(* Schneider Machine Expert - Basic project m200-cpp EXPERIMENTAL, file version 3.0.0.0 *)
(* ProjectInformations: Name=New project *)

HARDWARE
  Cpu 0: TM200CE40T
  EthernetConfiguration: NetworkName=M200, IpAllocationMode=FixedAddress, IpAddress=0.0.0.0, SubnetMask=0.0.0.0
  SerialLineConfiguration: Baud=Baud19200, Parity=ParityEven, DataBits=DataBits8, StopBits=StopBits1, PhysicalMedium=PhysicalMediumRs485, TransmissionMode=TransmissionModeModbusRtu, SlaveId=1, Addressing=SlaveAddressing
  MastTask: UsePeriodScanMode=false, PeriodScan=100
  FastTask: Period=255
  CpuBehavior: StartingMode=StartAsPreviousState, AutoSaveRamOnEeprom=true, WatchdogPeriod=250

SYMBOLS  (address, symbol, comment, settings)
  %S13      SB_FIRSTRUN  "Indicates the first controller cycle in RUN mode"
  %R0         [Type=Fifo]
  %M0       compiler_reused_M0_0
  %M1       compiler_reused_M1_1
  %M2       compiler_reused_M2_2
  %M3       compiler_reused_M3_3

POU Generated C++ - EXPERIMENTAL
  (* SectionNumber=0 *)

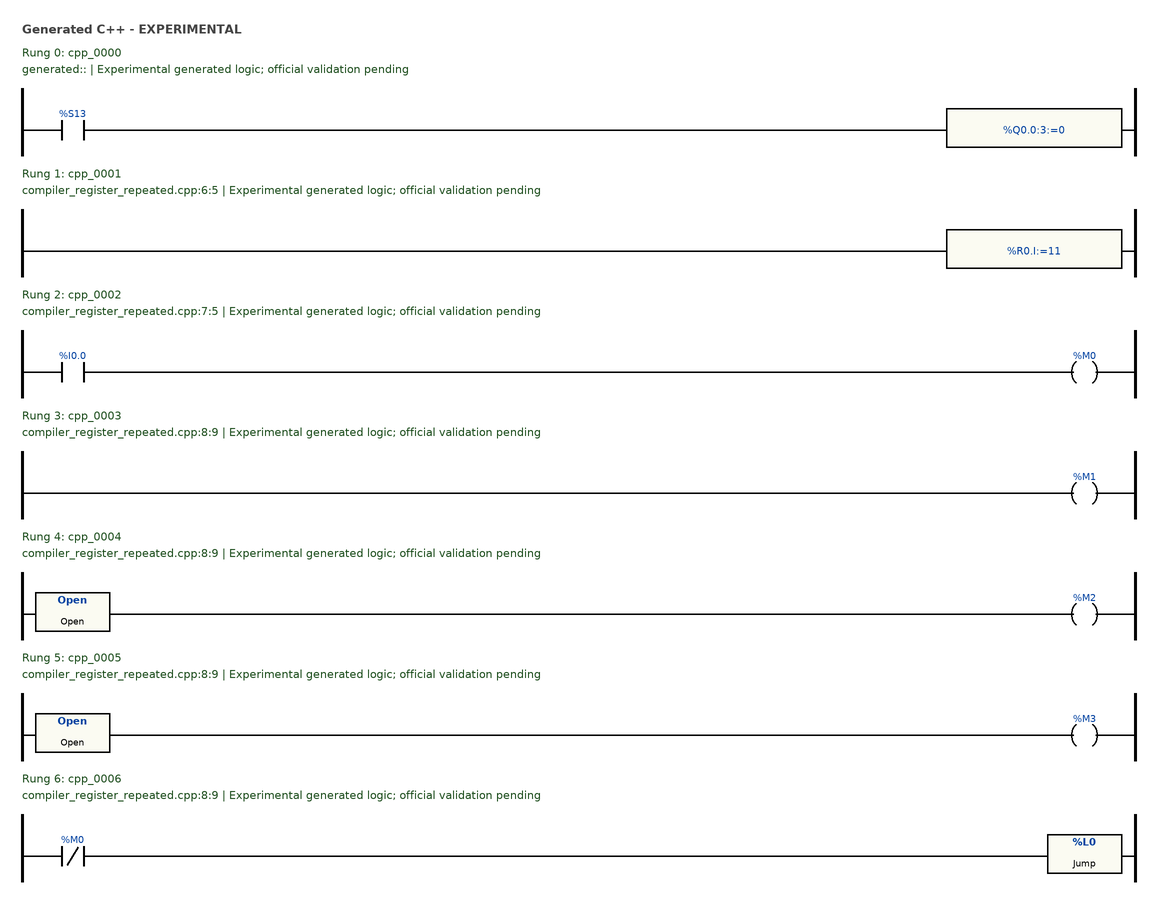

// Rung 0: cpp_0000
// generated:: | Experimental generated logic; official validation pending
  LD %S13                 (* SB_FIRSTRUN *)
  [%Q0.0:3:=0]
  // as ST:
  //   IF SB_FIRSTRUN THEN %Q0.0:3:=0; END_IF;

// Rung 1: cpp_0001
// compiler_register_repeated.cpp:6:5 | Experimental generated logic; official validation pending
  LD 1
  [%R0.I:=11]
  // as ST:
  //   %R0.I:=11;

// Rung 2: cpp_0002
// compiler_register_repeated.cpp:7:5 | Experimental generated logic; official validation pending
  LD %I0.0
  ST %M0                  (* compiler_reused_M0_0 *)
  // as ST:
  //   compiler_reused_M0_0 := %I0.0;

// Rung 3: cpp_0003
// compiler_register_repeated.cpp:8:9 | Experimental generated logic; official validation pending
  LD 1
  ST %M1                  (* compiler_reused_M1_1 *)
  // as ST:
  //   compiler_reused_M1_1 := TRUE;

// Rung 4: cpp_0004
// compiler_register_repeated.cpp:8:9 | Experimental generated logic; official validation pending
  LD 0
  ST %M2                  (* compiler_reused_M2_2 *)
  // as ST:
  //   compiler_reused_M2_2 := FALSE;

// Rung 5: cpp_0005
// compiler_register_repeated.cpp:8:9 | Experimental generated logic; official validation pending
  LD 0
  ST %M3                  (* compiler_reused_M3_3 *)
  // as ST:
  //   compiler_reused_M3_3 := FALSE;

// Rung 6: cpp_0006
// compiler_register_repeated.cpp:8:9 | Experimental generated logic; official validation pending
  LDN %M0                 (* compiler_reused_M0_0 *)
  JMPC %L0
  // as ST:
  //   IF NOT compiler_reused_M0_0 THEN JMP %L0; END_IF;

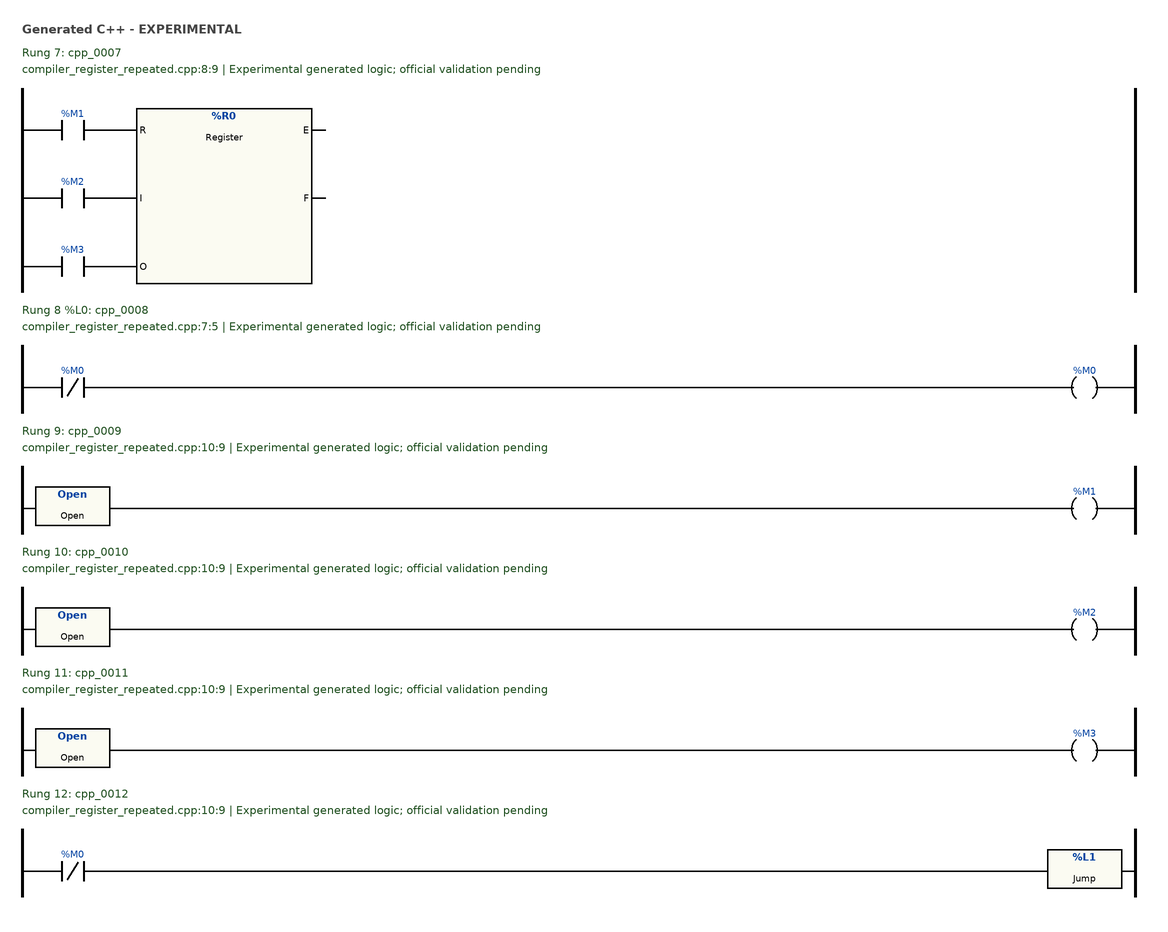

// Rung 7: cpp_0007
// compiler_register_repeated.cpp:8:9 | Experimental generated logic; official validation pending
  BLK %R0
  LD %M1                  (* compiler_reused_M1_1 *)
  R
  LD %M2                  (* compiler_reused_M2_2 *)
  I
  LD %M3                  (* compiler_reused_M3_3 *)
  O
  END_BLK
  // as ST:
  //   %R0(R := compiler_reused_M1_1, I := compiler_reused_M2_2, O := compiler_reused_M3_3);

// Rung 8 %L0: cpp_0008
// compiler_register_repeated.cpp:7:5 | Experimental generated logic; official validation pending
  %L0:
  LDN %M0                 (* compiler_reused_M0_0 *)
  ST %M0                  (* compiler_reused_M0_0 *)
  // as ST:
  //   %L0:
  //   compiler_reused_M0_0 := NOT compiler_reused_M0_0;

// Rung 9: cpp_0009
// compiler_register_repeated.cpp:10:9 | Experimental generated logic; official validation pending
  LD 0
  ST %M1                  (* compiler_reused_M1_1 *)
  // as ST:
  //   compiler_reused_M1_1 := FALSE;

// Rung 10: cpp_0010
// compiler_register_repeated.cpp:10:9 | Experimental generated logic; official validation pending
  LD 0
  ST %M2                  (* compiler_reused_M2_2 *)
  // as ST:
  //   compiler_reused_M2_2 := FALSE;

// Rung 11: cpp_0011
// compiler_register_repeated.cpp:10:9 | Experimental generated logic; official validation pending
  LD 0
  ST %M3                  (* compiler_reused_M3_3 *)
  // as ST:
  //   compiler_reused_M3_3 := FALSE;

// Rung 12: cpp_0012
// compiler_register_repeated.cpp:10:9 | Experimental generated logic; official validation pending
  LDN %M0                 (* compiler_reused_M0_0 *)
  JMPC %L1
  // as ST:
  //   IF NOT compiler_reused_M0_0 THEN JMP %L1; END_IF;

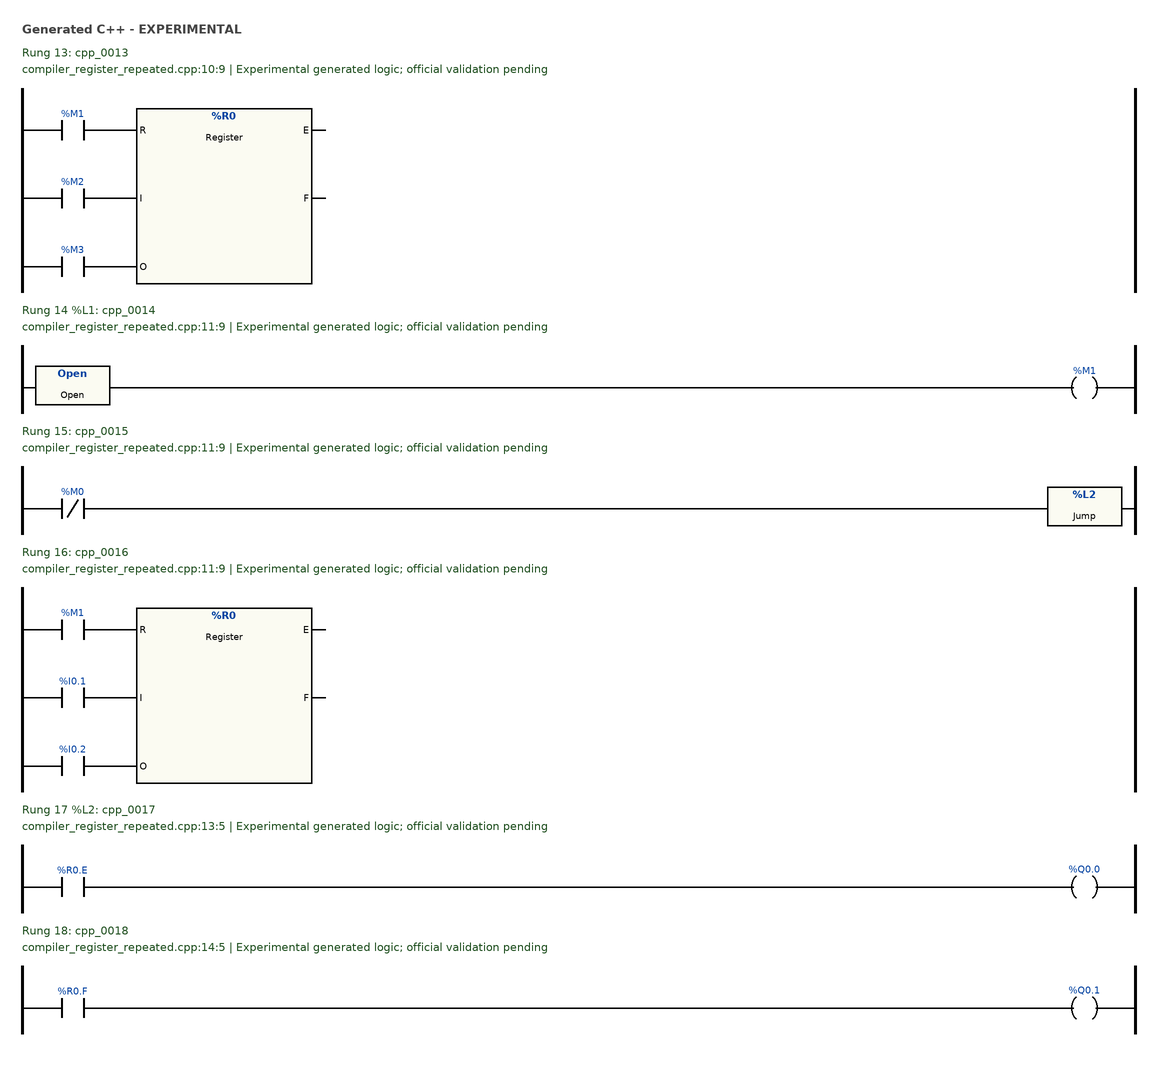

// Rung 13: cpp_0013
// compiler_register_repeated.cpp:10:9 | Experimental generated logic; official validation pending
  BLK %R0
  LD %M1                  (* compiler_reused_M1_1 *)
  R
  LD %M2                  (* compiler_reused_M2_2 *)
  I
  LD %M3                  (* compiler_reused_M3_3 *)
  O
  END_BLK
  // as ST:
  //   %R0(R := compiler_reused_M1_1, I := compiler_reused_M2_2, O := compiler_reused_M3_3);

// Rung 14 %L1: cpp_0014
// compiler_register_repeated.cpp:11:9 | Experimental generated logic; official validation pending
  %L1:
  LD 0
  ST %M1                  (* compiler_reused_M1_1 *)
  // as ST:
  //   %L1:
  //   compiler_reused_M1_1 := FALSE;

// Rung 15: cpp_0015
// compiler_register_repeated.cpp:11:9 | Experimental generated logic; official validation pending
  LDN %M0                 (* compiler_reused_M0_0 *)
  JMPC %L2
  // as ST:
  //   IF NOT compiler_reused_M0_0 THEN JMP %L2; END_IF;

// Rung 16: cpp_0016
// compiler_register_repeated.cpp:11:9 | Experimental generated logic; official validation pending
  BLK %R0
  LD %M1                  (* compiler_reused_M1_1 *)
  R
  LD %I0.1
  I
  LD %I0.2
  O
  END_BLK
  // as ST:
  //   %R0(R := compiler_reused_M1_1, I := %I0.1, O := %I0.2);

// Rung 17 %L2: cpp_0017
// compiler_register_repeated.cpp:13:5 | Experimental generated logic; official validation pending
  %L2:
  LD %R0.E
  ST %Q0.0
  // as ST:
  //   %L2:
  //   %Q0.0 := %R0.E;

// Rung 18: cpp_0018
// compiler_register_repeated.cpp:14:5 | Experimental generated logic; official validation pending
  LD %R0.F
  ST %Q0.1
  // as ST:
  //   %Q0.1 := %R0.F;

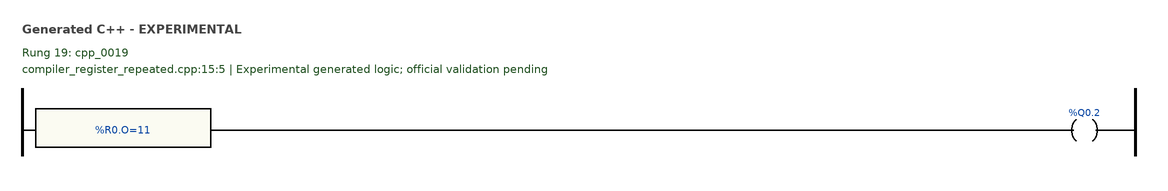

// Rung 19: cpp_0019
// compiler_register_repeated.cpp:15:5 | Experimental generated logic; official validation pending
  LD [%R0.O=11]
  ST %Q0.2
  // as ST:
  //   %Q0.2 := %R0.O=11;
